TYPE ST_PolarIIChamber_CupLiftServiceParam :
STRUCT
	JogPositive : ST_EmptyServiceParam;
	JogNegative : ST_EmptyServiceParam;
	IncrementalJog : ST_PolarIIChamber_LinearPositionParam;
	DecoupleStop : ST_EmptyServiceParam; // Speed, acceleration and deceleration are ECIDs.
	TopPos : ST_EmptyServiceParam;
	MiddlePos : ST_EmptyServiceParam;
	DownPos : ST_EmptyServiceParam;
END_STRUCT
END_TYPE

(* stored: Version 1.1.0.1, ProductVersion 3.1.4026.18
   DUT ST_PolarIIChamber_CupLiftServiceParam: Id {14000000-0000-0000-0000-000000000038} *)
